{attribute 'qualified_only'}
{attribute 'strict'}
{attribute 'to_string'}
TYPE E_Pump_List :
(
	eNotSelected := 0,
	P1001,
	P3001,
	P3002,
	P4001, //Line Color
	P4002, //CIP Color return
	TB0001,
	PP1002,
	PP1003,
	AG3001,
	AG3002,
	AG4001,
	AG4002,
	
	
	last
);
END_TYPE

(* stored: Version 1.1.0.1, ProductVersion 3.1.4024.13
   DUT E_Pump_List: Id {3ca80a79-00b9-4189-9306-867b9112375f} *)
